TYPE ST_HallOutputs :
STRUCT
    bOuterSpotsRelay : BOOL;
    bMiddleSpotRelay : BOOL;
END_STRUCT
END_TYPE

(* stored: Version 1.1.0.1
   DUT ST_HallOutputs: Id {6f05352e-02a2-45c4-9a58-d8076f2c820f} *)
